FUNCTION_BLOCK maximum2
VAR_INPUT
	x: ARRAY[0..243] OF LREAL;
	y: LREAL;
END_VAR
VAR_OUTPUT
	ex: ARRAY[0..243] OF LREAL;
END_VAR
VAR
	k: DINT;
END_VAR



FOR k := 0 TO 243 DO 
    ex[k] := MAX(x[k], y);
END_FOR;

END_FUNCTION_BLOCK

(* stored: Version 1.1.0.1, ProductVersion 3.1.4024.9
   POU maximum2: Id {ef7fbf74-8e70-4b36-b221-9f89e46cc15e}, SpecialFunc None *)
